(* IEC 61131-3 sources: rusty/tests/lit/single/type_promotion/bit_string/division, 6 files *)

(* ---- by_negative_literal.st ---- *)
// RUN: %COMPILE %s && %RUN | %CHECK %s
// XFAIL: *
// A negative literal next to a DWORD makes the division signed in 32 bits, and next to an LWORD it is read as unsigned.
FUNCTION main : DINT
    VAR
        dwmax : DWORD := 16#FFFF_FFFF;
        lw5 : LWORD := 16#5;
        r : LINT;
    END_VAR

    r := dwmax / -2;
    printf('DWORD max / -2 = %lld$N', r);                   // CHECK: DWORD max / -2 = -2147483647
    r := lw5 / -2;
    printf('LWORD 5 / -2 = %lld$N', r);                     // CHECK-NEXT: LWORD 5 / -2 = -2
END_FUNCTION

(* ---- byte_word_variables.st ---- *)
// RUN: %COMPILE %s && %RUN | %CHECK %s
// Two BYTE or WORD operands keep their own width, and their division and MOD are unsigned.
FUNCTION main : DINT
    VAR
        b : BYTE := 16#FF;
        b2 : BYTE := 16#02;
        b7 : BYTE := 16#07;
        w : WORD := 16#FFFF;
        w2 : WORD := 16#0002;
        w7 : WORD := 16#0007;
        rb : BYTE;
        rw : WORD;
    END_VAR

    rb := b / b2;
    printf('BYTE 16#FF / 2 = %u$N', rb);                    // CHECK: BYTE 16#FF / 2 = 127
    rb := b MOD b7;
    printf('BYTE 16#FF MOD 7 = %u$N', rb);                  // CHECK-NEXT: BYTE 16#FF MOD 7 = 3
    rw := w / w2;
    printf('WORD 16#FFFF / 2 = %u$N', rw);                  // CHECK-NEXT: WORD 16#FFFF / 2 = 32767
    rw := w MOD w7;
    printf('WORD 16#FFFF MOD 7 = %u$N', rw);                // CHECK-NEXT: WORD 16#FFFF MOD 7 = 1
END_FUNCTION

(* ---- division_guards.st ---- *)
// RUN: %COMPILE %s && %RUN | %CHECK %s
// Bit string divisions whose result does not depend on the type of the literal.
FUNCTION main : DINT
    VAR
        w : DWORD := 16#FFFF_FFFF;
        w2 : DWORD := 16#2;
        lw : LWORD := 16#FFFF_FFFF_FFFF_FFFF;
        qw : DWORD;
        ql : ULINT;
    END_VAR

    qw := w / w2;
    printf('DWORD max / DWORD 2 = %u$N', qw);               // CHECK: DWORD max / DWORD 2 = 2147483647
    ql := lw / 2;
    printf('LWORD max / 2 = %llu$N', ql);                   // CHECK-NEXT: LWORD max / 2 = 9223372036854775807
END_FUNCTION

(* ---- dword_by_untyped_literal.st ---- *)
// RUN: %COMPILE %s && %RUN | %CHECK %s
// An untyped integer literal takes the type of a DWORD operand, so the division is unsigned.
FUNCTION main : DINT
    VAR
        w : DWORD := 16#FFFF_FFFF;
        q : DWORD;
    END_VAR

    q := w / 2;
    printf('DWORD 16#FFFF_FFFF / 2 = %u$N', q);             // CHECK: DWORD 16#FFFF_FFFF / 2 = 2147483647
    q := w / 16#10;
    printf('DWORD 16#FFFF_FFFF / 16#10 = %u$N', q);         // CHECK-NEXT: DWORD 16#FFFF_FFFF / 16#10 = 268435455
    q := w MOD 3;
    printf('DWORD 16#FFFF_FFFF MOD 3 = %u$N', q);           // CHECK-NEXT: DWORD 16#FFFF_FFFF MOD 3 = 0
    q := w MOD 16#100;
    printf('DWORD 16#FFFF_FFFF MOD 16#100 = %u$N', q);      // CHECK-NEXT: DWORD 16#FFFF_FFFF MOD 16#100 = 255
END_FUNCTION

(* ---- with_signed_operand.st ---- *)
// RUN: %COMPILE %s && %RUN | %CHECK %s
// XFAIL: *
// A signed operand next to a DWORD makes the division signed, and next to an LWORD the bit string is read as negative,
// so a bit string from the signed midpoint on gives a wrong quotient.
FUNCTION main : DINT
    VAR
        i5 : INT := 5;
        i2 : INT := 2;
        l2 : LINT := 2;
        dwmax : DWORD := 16#FFFF_FFFF;
        lwmax : LWORD := 16#FFFF_FFFF_FFFF_FFFF;
        r : LINT;
    END_VAR

    r := dwmax / i2;
    printf('DWORD max / INT 2 = %lld$N', r);                // CHECK: DWORD max / INT 2 = 2147483647
    r := i5 MOD dwmax;
    printf('INT 5 MOD DWORD max = %lld$N', r);              // CHECK-NEXT: INT 5 MOD DWORD max = 5
    r := lwmax / l2;
    printf('LWORD max / LINT 2 = %lld$N', r);               // CHECK-NEXT: LWORD max / LINT 2 = 9223372036854775807
END_FUNCTION

(* ---- literal_by_declaration_section.st ---- *)
// RUN: %COMPILE %s && %RUN | %CHECK %s
// A DWORD operand divided by an untyped literal stays DWORD, wherever the operand is declared.
VAR_GLOBAL
    g : DWORD := 16#FFFF_FFFF;
END_VAR

VAR_GLOBAL CONSTANT
    gc : DWORD := 16#FFFF_FFFF;
END_VAR

FUNCTION_BLOCK probe
    VAR_INPUT
        i : DWORD;
    END_VAR
    VAR_INPUT CONSTANT
        ic : DWORD := 16#FFFF_FFFF;
    END_VAR
    VAR_IN_OUT
        io : DWORD;
    END_VAR
    VAR_OUTPUT
        o : DWORD;
    END_VAR
    VAR CONSTANT
        c : DWORD := 16#FFFF_FFFF;
    END_VAR
    VAR_TEMP
        t : DWORD;
    END_VAR
    VAR
        q : ULINT;
    END_VAR

    o := 16#FFFF_FFFF;
    t := 16#FFFF_FFFF;
    q := i / 2;
    printf('VAR_INPUT / 2 = %llu$N', q);
    q := ic MOD 7;
    printf('VAR_INPUT CONSTANT MOD 7 = %llu$N', q);
    q := io / 2;
    printf('VAR_IN_OUT / 2 = %llu$N', q);
    q := io MOD 7;
    printf('VAR_IN_OUT MOD 7 = %llu$N', q);
    q := o / 2;
    printf('VAR_OUTPUT / 2 = %llu$N', q);
    q := c MOD 7;
    printf('VAR CONSTANT MOD 7 = %llu$N', q);
    q := t / 2;
    printf('VAR_TEMP / 2 = %llu$N', q);
    q := g MOD 7;
    printf('VAR_GLOBAL MOD 7 = %llu$N', q);
    q := gc / 2;
    printf('VAR_GLOBAL CONSTANT / 2 = %llu$N', q);
END_FUNCTION_BLOCK

FUNCTION main : DINT
    VAR
        inst : probe;
        v : DWORD := 16#FFFF_FFFF;
    END_VAR

    inst(i := 16#FFFF_FFFF, io := v);
    // CHECK: VAR_INPUT / 2 = 2147483647
    // CHECK-NEXT: VAR_INPUT CONSTANT MOD 7 = 3
    // CHECK-NEXT: VAR_IN_OUT / 2 = 2147483647
    // CHECK-NEXT: VAR_IN_OUT MOD 7 = 3
    // CHECK-NEXT: VAR_OUTPUT / 2 = 2147483647
    // CHECK-NEXT: VAR CONSTANT MOD 7 = 3
    // CHECK-NEXT: VAR_TEMP / 2 = 2147483647
    // CHECK-NEXT: VAR_GLOBAL MOD 7 = 3
    // CHECK-NEXT: VAR_GLOBAL CONSTANT / 2 = 2147483647
END_FUNCTION
